// TIA Portal V20 export
Screen "Pop-up_NutRunner"  395x450
  ScreenItem "Robot Name" at 2,2 size 393x48  Type=HmiIOField
  ScreenItem "Background" at -1,49 size 395x400  Type=HmiRectangle
  ScreenItem "Cancel Mode" at 315,4 size 76x42  Type=HmiButton
  ScreenItem "矩形_4" at 29,71 size 324x285  Type=HmiRectangle
  ScreenItem "Text Field In Auto On_9" at 41,107 size 148x21  Type=HmiTextBox
  ScreenItem "Text Field Home Position_17" at 41,131 size 148x21  Type=HmiTextBox
  ScreenItem "Text field Robot Status_5" at 27,72 size 328x30  Type=HmiTextBox
  ScreenItem "Text Field Manual_17" at 41,275 size 148x21  Type=HmiTextBox
  ScreenItem "Text Field System Ready_9" at 41,155 size 148x21  Type=HmiTextBox
  ScreenItem "Text Field Motor On_9" at 41,179 size 148x21  Type=HmiTextBox
  ScreenItem "Text Field In Cycle_9" at 41,203 size 148x21  Type=HmiTextBox
  ScreenItem "Text Field Cycle On_17" at 41,227 size 148x21  Type=HmiTextBox
  ScreenItem "Text Field On Path_17" at 41,251 size 148x21  Type=HmiTextBox
  ScreenItem "Text Field Home Position_18" at 196,107 size 148x21  Type=HmiTextBox
  ScreenItem "Text Filed E- Stop_18" at 196,251 size 148x21  Type=HmiTextBox
  ScreenItem "Text Field Manual_18" at 196,179 size 148x21  Type=HmiTextBox
  ScreenItem "Text Field Cycle On_18" at 196,131 size 148x21  Type=HmiTextBox
  ScreenItem "Text Field On Path_18" at 196,155 size 148x21  Type=HmiTextBox
  ScreenItem "Text Field Tryout Mode_18" at 196,203 size 148x21  Type=HmiTextBox
  ScreenItem "Text Field Stop_18" at 196,227 size 148x21  Type=HmiTextBox
  ScreenItem "Text Field In Auto On_10" at 196,275 size 148x21  Type=HmiTextBox
